(* IEC 61131-3 sources: ConveyorControl-with-PLC/4E_Gruppe1_Graf_Projekt1/Network/net0, 1 file *)

(* ---- ONE_net0_Table.st ---- *)
#define OBJECTS_CONFIG

FUNCTION GLOBAL TAB ONE_net0
-1$UINT, 0$UINT,
0$UINT, 0$UINT,

1$UDINT,
TO_UDINT(1869306653), "Abschluss", 0$UINT, 0$UINT, 1$UINT,

_NO_ATTR, TO_UDINT(3770017845), "ABSCHLUSS1",

//Internal connections
0$UDINT,
0$UDINT,
0$UDINT,
0$UDINT,

//Initialization values
0$UDINT,
0$UDINT,

//Symbolic initialization values
0$UDINT,
0$UDINT,

//Initialization of string values
0$UDINT,
0$UDINT,

//Configuration of tasks (RealTime, Cyclic, Background)
0$UDINT,
0$UDINT,

0$UDINT,
1$UDINT,
TO_UDINT(0), (10)$UDINT, 4194303$DINT, 	//ABSCHLUSS1

0$UDINT,
0$UDINT,

//External connections
0$UDINT,
2$UDINT,
TO_UDINT(0), "MTR_speed", C_DIR, TO_UDINT(3059689190), "_DriveAxis1","SetSpeed",
TO_UDINT(0), "MTR_enable", C_DIR, TO_UDINT(3059689190), "_DriveAxis1","AxEnable",

//Magic internal connections
0$UDINT,
0$UDINT,

//Configuration of timeslots of tasks (RealTime, Cyclic)
#ifdef __LSLLDR_TIMESLOTS__
0$UDINT,
0$UDINT,

0$UDINT,
0$UDINT,

#endif //__LSLLDR_TIMESLOTS__

//MultiMaster connections
#ifdef __LSLLDR_MULTIMASTER__
0$UDINT,
0$UDINT,
#endif //__LSLLDR_MULTIMASTER__

END_FUNCTION
